Fanuc KAREL source: kc00020.KL

-- PROVISIONAL review KL for V940-1; original PC SHA256 14829a7e77f99700fe4f8d06ca3b539092cd9298767d85edddeee6c41b865ab6
-- Incomplete behavior may be omitted. Consult companion uncertainty JSON. Do not deploy.
PROGRAM KC00020
%NOLOCKGROUP
BEGIN
  -- V9_ZERO_TABLE_METADATA_HINT layout=0002_ascii; no indexed target words; source/name/runtime held
  -- UNRESOLVED_PC offsets 5-12; opcodes 27,27,27,9C,31
  -- UNRESOLVED_PC offsets 17-21; opcodes 7F
END KC00020
